Fanuc KAREL source: kc00015.KL

-- PROVISIONAL review KL for V770-1; original PC SHA256 b39ce65b06cf34b9e1acdde65f25b0b73c71a293f82b67b64d55c9554fb3d7bd
-- Incomplete behavior may be omitted. Consult companion uncertainty JSON. Do not deploy.
PROGRAM KC00015
%NOLOCKGROUP
BEGIN
  -- UNRESOLVED_PC offsets 5-12; opcodes 9D,23
  -- UNRESOLVED_PC offsets 17-47; opcodes 27,22,22,27,9D,31,7E,4A
  -- UNRESOLVED_PC offsets 52-56; opcodes 7F
END KC00015
